(* IEC 61131-3 sources: STAR-PLC-Agent/results/raw/compiler_smoke_2026-11-10T120847007597+0000/repaired, 1 file *)

(* ---- FB_Task.st ---- *)
FUNCTION_BLOCK FB_Task
VAR_INPUT
 Start : BOOL;
 Stop : BOOL;
END_VAR
VAR_OUTPUT
 Run : BOOL := FALSE;
END_VAR

IF Stop THEN
 Run := FALSE;
ELSIF Start THEN
 Run := TRUE;
END_IF;
END_FUNCTION_BLOCK
